TYPE ST_PolarIIChamber_FlowCalibrationParam :
STRUCT
	ArmIndex : UINT; // 1..4
	ArmNozzleIndex : UINT; // 1..3
	TestTime : TIME;
END_STRUCT
END_TYPE

(* stored: Version 1.1.0.1, ProductVersion 3.1.4026.18
   DUT ST_PolarIIChamber_FlowCalibrationParam: Id {14000000-0000-0000-0000-000000000018} *)
